(* PLC project probe, plc-portfolio cds2astra probe 0.1.0 *)
(* stored: creationDateTime 2026-10-20T00:00:00, modificationDateTime 2026-10-20T00:00:00 *)

{attribute 'symbol' := 'read'}
PROGRAM PRG_P3
VAR
    fbHyst : HYSTERESIS;
END_VAR

            fbHyst(IN := 50, HIGH := 80, LOW := 20);
          
END_PROGRAM
